FUNCTION_BLOCK FB_CompD_1
(*
Function block used to calculate differential typ.

Constructor: 		Patryk Panylo
Company:		E. Riexinger GmbH
Date:			03.06.2014
Version:			1.00

Date:			Revision:		Who:				Comment
dd.mm.yyyy		x.xx			Initials			comment

*)

VAR_INPUT
	(* Enummerations *)

	(* Variables *)
	bEnable								:BOOL := TRUE;					(* Enable FB *)
	lrInSignal								:LREAL;							(* Input signal *)
	lrDifferentialValue						:LREAL := 1.0;						(* Differential value *)
	lrTaskCycle							:LREAL := 1.0; 					(* Cycle time *)


	(* References *)

	(* Interfaces *)

	(* Instances *)

END_VAR
VAR_OUTPUT
	(* Enummerations *)

	(* Variables *)
	lrOutSignal							:LREAL;							(* Output signal *)

	(* References *)

	(* Interfaces *)

	(* Instances *)
END_VAR
VAR
	(* Enummerations *)

	(* Variables *)
	bFirstTime							:BOOL;							(* First cycle *)

	(* References *)

	(* Interfaces *)

	(* Instances *)
	fbDifferential								:FB_Differential;

END_VAR

IF NOT bEnable
THEN

	fbDifferential(
		bEnable := FALSE,
		lrInSignal := lrInSignal,
		lrDifferentialValue := lrDifferentialValue,
		lrTaskCycle := lrTaskCycle,
		lrOutSignal => lrOutSignal
	);

	bFirstTime := FALSE;
	RETURN;
END_IF

IF NOT bFirstTime
THEN
	bFirstTime := TRUE;
END_IF

A_CalcDifferential();

ACTION A_CalcDifferential:

fbDifferential(
	bEnable := TRUE,
	lrInSignal := lrInSignal,
	lrDifferentialValue := lrDifferentialValue,
	lrTaskCycle := lrTaskCycle,
	lrOutSignal => lrOutSignal
);
END_ACTION

END_FUNCTION_BLOCK

(* stored: Version 1.1.0.1, ProductVersion 3.1.4024.15
   POU FB_CompD_1: Id {a3b087de-bbf9-4bd9-a13f-619c47a72b89}, SpecialFunc None
   Action A_CalcDifferential: Id {0b41511e-c548-4d03-b026-e0557aba418d} *)
